// TIA Portal V17 export
// export: Created 2026-11-08T05:50:27.715777Z, ExportSetting WithDefaults, DisplayName Totally Integrated Automation Portal, DisplayVersion V17, DisplayName TIA Portal Openness, DisplayVersion V17, DisplayName TIA Portal Version Control Interface, DisplayVersion V17, DisplayName STEP 7 Professional, DisplayVersion V17, DisplayName STEP 7 Safety, DisplayVersion V17, DisplayName WinCC Professional, DisplayVersion V17
DATA_BLOCK "DB_Mando"   // DB2
VERSION : 0.1
// stored: AutoNumber true, DBAccessibleFromOPCUA true, InstanceOfName FB_Mando_Motor, InstanceOfType FB
"FB_Mando_Motor"
   // VAR_INPUT
   //    PB_Marcha : Bool;
   //    PB_Paro : Bool;
   //    Termico_Falla : Bool;
   //    HMI_Marcha : Bool;
   //    HMI_Paro : Bool;
   //    HMI_Reset : Bool;
   // END_VAR
   // VAR_OUTPUT
   //    Marcha : Bool;
   //    Paro : Bool;
   //    Termico_OK : Bool;
   //    Reset : Bool;
   // END_VAR
   // VAR
   //    T_Reset : TON_TIME;
   //    Reset_Mantenido : Bool;
   // END_VAR
BEGIN
END_DATA_BLOCK
